FUNCTION_BLOCK AckLedControl (* Composite Function Block Type *)
  (* Standard: 61499-2 *)
  (* Version 0.0, 10/19/2026, macie, Schneider Electric, template *)
  PACKAGE Main;
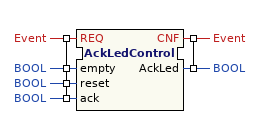
  EVENT_INPUT
    REQ WITH empty, reset, ack; (* Normal Execution Request *)
  END_EVENT
  EVENT_OUTPUT
    CNF WITH AckLed; (* Execution Confirmation *)
  END_EVENT
  VAR_INPUT
    empty : BOOL; (* Input event qualifier *)
    reset : BOOL;
    ack : BOOL;
  END_VAR
  VAR_OUTPUT
    AckLed : BOOL; (* Output event qualifier *)
  END_VAR
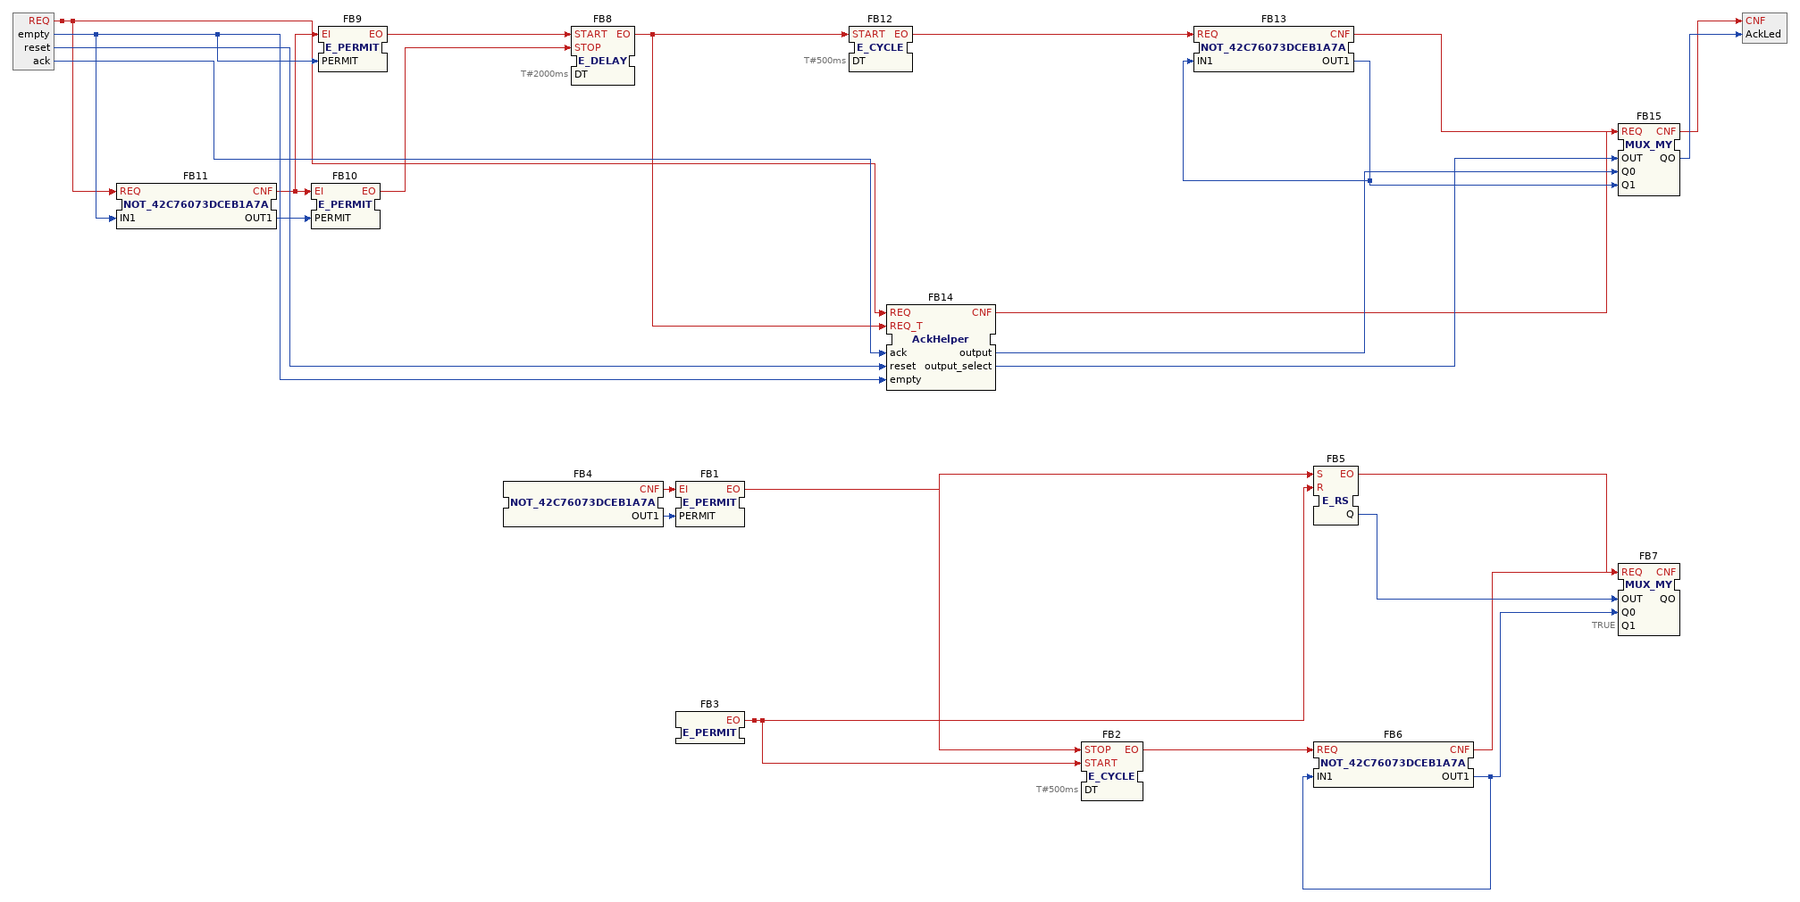
  FBS
    FB1 : E_PERMIT;
    FB2 : E_CYCLE(DT := T#500ms);
    FB3 : E_PERMIT;
    FB4 : NOT_42C76073DCEB1A7A; {SET_ATTRIBUTE(Configuration.GenericFBType.InterfaceParams, Runtime.Standard#CNT:=1;OUT${CNT$}:BOOL)}
    FB6 : NOT_42C76073DCEB1A7A; {SET_ATTRIBUTE(Configuration.GenericFBType.InterfaceParams, Runtime.Standard#CNT:=1;OUT${CNT$}:BOOL)}
    FB5 : E_RS;
    FB7 : MUX_MY(Q1 := TRUE);
    FB8 : E_DELAY(DT := T#2000ms);
    FB9 : E_PERMIT;
    FB10 : E_PERMIT;
    FB11 : NOT_42C76073DCEB1A7A; {SET_ATTRIBUTE(Configuration.GenericFBType.InterfaceParams, Runtime.Standard#CNT:=1;OUT${CNT$}:BOOL)}
    FB12 : E_CYCLE(DT := T#500ms);
    FB13 : NOT_42C76073DCEB1A7A; {SET_ATTRIBUTE(Configuration.GenericFBType.InterfaceParams, Runtime.Standard#CNT:=1;OUT${CNT$}:BOOL)}
    FB15 : MUX_MY;
    FB14 : AckHelper;
  END_FBS
  EVENT_CONNECTIONS
    FB4.CNF TO FB1.EI;
    FB2.EO TO FB6.REQ;
    FB1.EO TO FB5.S;
    FB3.EO TO FB5.R;
    FB1.EO TO FB2.STOP;
    FB3.EO TO FB2.START;
    FB6.CNF TO FB7.REQ;
    FB5.EO TO FB7.REQ;
    REQ TO FB11.REQ;
    FB11.CNF TO FB10.EI;
    FB11.CNF TO FB9.EI;
    FB9.EO TO FB8.START;
    FB10.EO TO FB8.STOP;
    FB8.EO TO FB12.START;
    FB12.EO TO FB13.REQ;
    FB15.CNF TO CNF;
    FB13.CNF TO FB15.REQ;
    FB8.EO TO FB14.REQ_T;
    REQ TO FB14.REQ;
    FB14.CNF TO FB15.REQ;
  END_CONNECTIONS
  DATA_CONNECTIONS
    FB4.OUT1 TO FB1.PERMIT;
    FB6.OUT1 TO FB6.IN1;
    FB5.Q TO FB7.OUT;
    FB6.OUT1 TO FB7.Q0;
    empty TO FB9.PERMIT;
    FB11.OUT1 TO FB10.PERMIT;
    empty TO FB11.IN1;
    FB13.OUT1 TO FB13.IN1;
    FB15.QO TO AckLed;
    FB13.OUT1 TO FB15.Q1;
    ack TO FB14.ack;
    reset TO FB14.reset;
    FB14.output TO FB15.Q0;
    FB14.output_select TO FB15.OUT;
    empty TO FB14.empty;
  END_CONNECTIONS
END_FUNCTION_BLOCK
